Universal Robots URScript: T008_qwen2.5-coder_32b_baseline_rep1.urscript

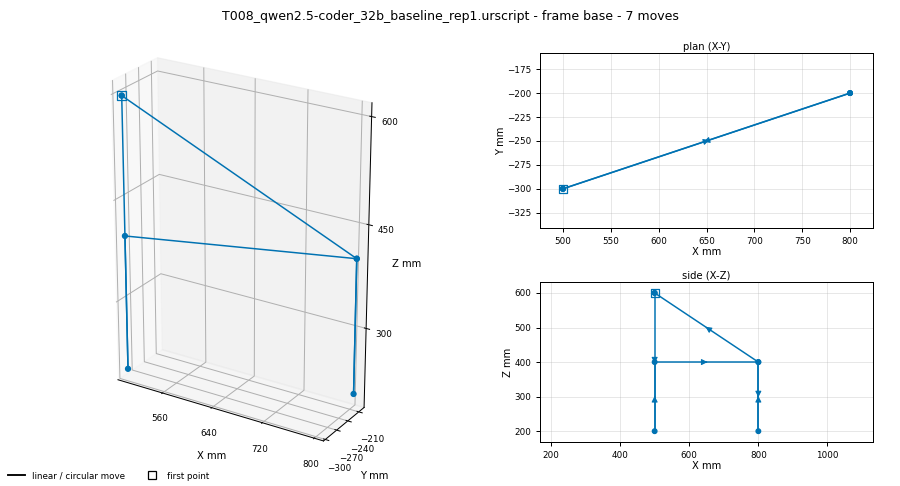
[picture p0: tool path of T008_qwen2.5-coder_32b_baseline_rep1.urscript in frame base, 7 of 9 moves have a stored position in this frame; points joined in program order, loops and branches not executed]
def depalletize_heavy_boxes():
    # Move to Home position
    movej(get_inverse_kin([0, -90, 90, -90, 90, 0]), a=1.4, v=1.2)

    # Move above pallet
    movel(p[0.5, -0.3, 0.6, 3.14, 0, 0], a=1.2, v=1.0)

    # Descend to top layer of pallet
    movel(p[0.5, -0.3, 0.2, 3.14, 0, 0], a=0.8, v=0.6)

    # Lift box from pallet
    movel(p[0.5, -0.3, 0.4, 3.14, 0, 0], a=0.7, v=0.5)

    # Transit to conveyor
    movel(p[0.8, -0.2, 0.4, 3.14, 0, 0], a=1.0, v=0.9)

    # Place box on conveyor
    movel(p[0.8, -0.2, 0.2, 3.14, 0, 0], a=0.7, v=0.5)

    # Lift TCP from conveyor
    movel(p[0.8, -0.2, 0.4, 3.14, 0, 0], a=0.7, v=0.5)

    # Return above pallet for next box
    movel(p[0.5, -0.3, 0.6, 3.14, 0, 0], a=1.2, v=1.0)

    # Move to Home position
    movej(get_inverse_kin([0, -90, 90, -90, 90, 0]), a=1.4, v=1.2)
end

depalletize_heavy_boxes()
